Fanuc KAREL source: KT00608.KL

PROGRAM KT00608
%NOLOCKGROUP
VAR
  R1: REAL
  R2: REAL
  OUT: REAL
BEGIN
  R1 = 2.0
  R2 = 3.0
  R1 = 2.0
  R2 = 3.0
  OUT = NOT R1
END KT00608
